Fanuc KAREL source: KA00055.KL

PROGRAM KA00055
%NOLOCKGROUP
VAR
  SRC: POSITION
  DST: XYZWPREXT
BEGIN
  DST = SRC
END KA00055
